Fanuc KAREL source: kb00023.compact.KL

PROGRAM KB00023
%STACKSIZE=65535
%PRIORITY=65535
%NOLOCKGROUP
VAR
P1 : INTEGER
P2 : INTEGER
BEGIN
P1=1
P2=1
CLOSE_TPE(P1,P2)
END KB00023
